FUNCTION_BLOCK PI_Function_Block
VAR_INPUT
    Setpoint :REAL := 54;
    Actual: REAL;
	Bias: REAL := 40;
    Kp :REAL := 20;
    Ti :REAL := 40;
    Td :REAL := 0;
    Ts :REAL := 0.01;
    N :REAL := 1;
    OutMax :REAL := 100;
    OutMin :REAL := 0;
    bEuler :BOOL := FALSE;
	bEnable :BOOL;
END_VAR

VAR_OUTPUT
    Output :REAL;
    Error :REAL;
END_VAR

VAR
    PrevError :REAL;
    Integ :REAL;
    Deriv :REAL;
    dInteg :REAL;
    Tf :REAL;
    DerivRaw :REAL;
    Unsat :REAL;
END_VAR

Error := Actual - Setpoint;

IF NOT bEnable THEN
	Integ := 0.0;
	dInteg := 0.0;
	Output := Main.Level_Valve_2_Percentage;
	RETURN;
END_IF

IF Ti > 0.0 THEN
    IF bEuler THEN
    dInteg := Ts / Ti * Error;
ELSE
    dInteg := Ts / Ti * (Error + PrevError) / 2;
END_IF
ELSE
    dInteg := 0.0;
    Integ := 0.0;
END_IF

IF N > 0.0 THEN
    Tf := Td / N;
ELSE
    Tf := 0.0;
END_IF

DerivRaw := Td * (Error - PrevError) / Ts;
Deriv := (Tf * Deriv + Ts * DerivRaw)
/ (Tf + Ts);

Unsat := Kp * (Error + Integ + dInteg + Deriv) + Bias;

IF (Unsat > OutMax AND dInteg > 0) OR
(Unsat < OutMin AND dInteg < 0) THEN
dInteg := 0; // anti-windup
END_IF
Integ := Integ + dInteg;

Output := Kp * (Error + Integ + Deriv) + Bias;
IF Output > OutMax THEN Output := OutMax; END_IF
IF Output < OutMin THEN Output := OutMin; END_IF

PrevError := Error;

END_FUNCTION_BLOCK

(* stored: Version 1.1.0.1, ProductVersion 3.1.4026.21
   POU PI_Function_Block: Id {efb42321-a56f-439b-a67e-f0f245e3bee1}, SpecialFunc None *)
